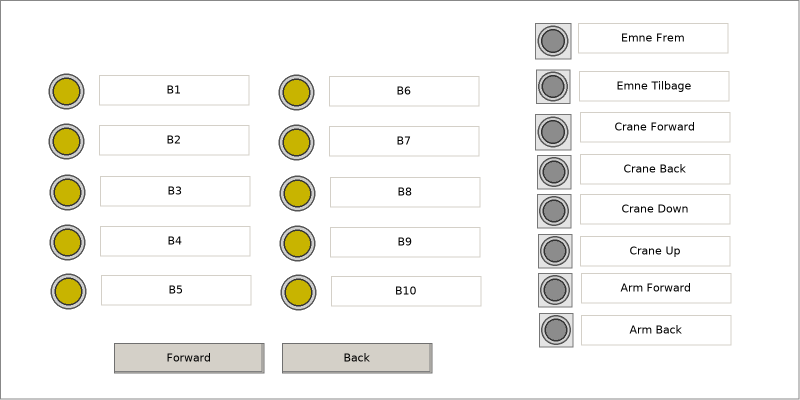
VISUALIZATION IO  // 800x400
    Lamp1 (46,71 41x41), variable: MAIN.B1, style: Lamp-Lamp1-Yellow
    Textfield (99,75 150x30), "B1"
    Textfield (99,125 150x30), "B2"
    Lamp1 (46,121 41x41), variable: MAIN.B2, style: Lamp-Lamp1-Yellow
    Lamp1 (47,172 41x41), variable: MAIN.B3, style: Lamp-Lamp1-Yellow
    Textfield (100,176 150x30), "B3"
    Textfield (100,226 150x30), "B4"
    Lamp1 (47,222 41x41), variable: MAIN.B4, style: Lamp-Lamp1-Yellow
    Lamp1 (48,271 41x41), variable: MAIN.B5, style: Lamp-Lamp1-Yellow
    Textfield (101,275 150x30), "B5"
    Lamp1 (276,72 41x41), variable: MAIN.B6, style: Lamp-Lamp1-Yellow
    Textfield (329,76 150x30), "B6"
    Textfield (329,126 150x30), "B7"
    Lamp1 (276,122 41x41), variable: MAIN.B7, style: Lamp-Lamp1-Yellow
    Lamp1 (277,173 41x41), variable: MAIN.B8, style: Lamp-Lamp1-Yellow
    Textfield (330,177 150x30), "B8"
    Textfield (330,227 150x30), "B9"
    Lamp1 (277,223 41x41), variable: MAIN.B9, style: Lamp-Lamp1-Yellow
    Lamp1 (278,272 41x41), variable: MAIN.B10, style: Lamp-Lamp1-Yellow
    Textfield (331,276 150x30), "B10"
    Textfield (579,71 150x30), "Emne Tilbage"
    PushSwitch (536,69 34x35), variable: MAIN.M1_Forward, behaviour: TAP, style: Switch-PushSwitch-Gray
    PushSwitch (535,23 36x36), variable: MAIN.M1_Back, behaviour: TAP, style: Switch-PushSwitch-Gray
    Textfield (578,23 150x30), "Emne Frem"
    Textfield (580,112 150x30), "Crane Forward"
    PushSwitch (535,114 36x36), variable: MAIN.M2_Forward, behaviour: TAP, style: Switch-PushSwitch-Gray
    PushSwitch (537,155 34x34), variable: MAIN.M2_Back, behaviour: TAP, style: Switch-PushSwitch-Gray
    Textfield (580,154 150x30), "Crane Back"
    Textfield (580,194 150x30), "Crane Down"
    PushSwitch (537,194 34x34), variable: MAIN.M3_Down, behaviour: TAP, style: Switch-PushSwitch-Gray
    PushSwitch (538,234 34x34), variable: MAIN.M3_Up, behaviour: TAP, style: Switch-PushSwitch-Gray
    Textfield (580,236 150x30), "Crane Up"
    Textfield (581,273 150x30), "Arm Forward"
    PushSwitch (538,273 34x34), variable: MAIN.M4_Forward, behaviour: TAP, style: Switch-PushSwitch-Gray
    PushSwitch (539,313 34x34), variable: MAIN.M4_Back, behaviour: TAP, style: Switch-PushSwitch-Gray
    Textfield (581,315 150x30), "Arm Back"
    Button (114,343 150x30), "Forward"
        tap MAIN.bJogForward
    Button (282,343 150x30), "Back"
        tap MAIN.bJogBackward
END_VISUALIZATION

(* stored: Version 1.1.0.1, ProductVersion 3.1.4024.12
   Visu IO: Id {8da2a5a5-256d-4ba0-861e-2393506b703d} *)
